FUNCTION_BLOCK TPBLOCK
VAR_INPUT
	in:BOOL;
	pt:TIME;
	
END_VAR
VAR_OUTPUT
	out:BOOL;
	et:TIME;
	
END_VAR
VAR
	tstarttime:TIME;
	bpulseact:BOOL;
	bprevin:BOOL;
	

END_VAR

IF in AND NOT bprevin AND NOT bpulseact THEN
	tstarttime:=TIME();
	bpulseact:=TRUE;
	out:=TRUE;
	et:=T#0MS;
	
END_IF
IF bpulseact THEN 
	et:=TIME()-tstarttime;
	IF et>= pt THEN 
		et:=pt;
		out:=FALSE;
		bpulseact:=FALSE;
	END_IF
ELSE
	IF NOT in THEN
		et:=T#0MS;
	END_IF
END_IF

END_FUNCTION_BLOCK

(* stored: Version 1.1.0.1, ProductVersion 3.1.4024.16
   POU TPBLOCK: Id {feedda1d-f846-4973-b3cb-fc5eb4e3d362}, SpecialFunc None *)
